(* IEC 61131-3 sources: trust-platform/conformance/cases/timers/cfm_timers_ton_sequence_001, 1 file *)

(* ---- program.st ---- *)
PROGRAM Main
VAR
    ton_fb : TON;
    in_ton : BOOL;
    q_ton : BOOL;
    et_ton : TIME;
END_VAR

ton_fb(IN := in_ton, PT := T#10ms, Q => q_ton, ET => et_ton);
END_PROGRAM
